(* IEC 61131-3 sources: BODAS-HelloWorld/st/bodas_rc18_12_40/plc_logic/application/02_easyconfig/easyconfig_import/bds_syspb_ec, 2 files *)

(* ---- bds_syspb_vrnt_te-bds_sysPb_vrnt_te.st ---- *)
(* --- Interface --- *)
///post build system variants information
{attribute 'qualified_only' := ''}
{attribute 'strict' := ''}
TYPE bds_sysPb_vrnt_te : (
		bds_sysPb_vrnt01_E := 0,
		bds_sysPb_maxNumVrnt_E
	) USINT;
END_TYPE

(* ---- bds_syspb_ec_gvl-bds_sysPb_ec_gvl.st ---- *)
(* --- Interface --- *)
{attribute 'qualified_only' := ''}
VAR_GLOBAL CONSTANT
	ml290rts_bs_HelloWorld : USINT := bds_sysPb_vrnt_te.bds_sysPb_vrnt01_E;
END_VAR
